(* IEC 61131-3 sources: JingjiangMoonbox/Application/Application/任务列表/Main_Task/套色调整/新算法/JIEOU, 8 files *)

(* ---- JIEOU10.st ---- *)
(*@CES
Name=JIEOU10
Type=FunctionBlock
TypeGuid=6f9dac99-8de1-4efc-8465-68ac443b7d08
Guid=2b28cbf0-4862-4f21-a282-23685e336d72
HasDeclaration=True
HasImplementation=True
*)
{DECLARATION}
FUNCTION JIEOU10 : REAL
VAR_INPUT
	i_rPI2_AND_JIEOU3_AND_JIEOU4:REAL;(*PI2和JIEOU3JIEOU4经过JIEOU8 Gc2Yk_K5_K6的输出/Gc2Uk_K5_K6输入*)
	i_rJIEOU5:REAL;(*U5经过JIEOU8 Gc2Yk_K3的输出/Gc2Uk_K4输入*)
	i_rJIEOU6:REAL;(*U6经过JIEOU9 Gc2Yk_K3的输出*)
	i_rJIEOU7:REAL;(*U7经过JIEOU9 Gc2_1的输出*)
	i_rJIEOU8:REAL;(*U8输出*)
	i_rJIEOU9:REAL;(*U9输出*)
	i_rPI10:REAL;(*PI10输出*)

	i_prU10: POINTER TO REAL;(*解耦后控制器8输出*)

(*
	i_rL:REAL;(*版周长mm*)
	i_rV:REAL;(*运行速度m/min*)
*)
	i_rTs:REAL;(*2024.6.29.135040修改为了输入@s*)
	i_rA:REAL;(*系统参数A*)
(*Gc1_1寄存器*)
	i_prGc1_1_Uk:POINTER TO ARRAY [1..ARC_DELAY_N_MAX] OF REAL;(*Gc1_1输入寄存器*)
	i_prGc1_1_Gc1_Yk:POINTER TO ARRAY [1..2] OF REAL;(*Gc1_1 Gc1输出寄存器*)
(*Gc2_1寄存器*)
	i_prGc2_1_Uk:POINTER TO ARRAY [1..ARC_DELAY_N_MAX] OF REAL;(*Gc2_1输入寄存器*)
	i_prGc2_1_Yk:POINTER TO ARRAY [1..2] OF REAL;(*Gc2_1输出寄存器*)

	i_prGc2_1_Gc1_Uk:POINTER TO ARRAY [1..2] OF REAL;(*Gc2_1 Gc1输入寄存器*)
	i_prGc2_1_Gc2_Yk:POINTER TO ARRAY [1..2] OF REAL;(*Gc2_1 Gc2输出寄存器*)

(*Gc2寄存器3*)
	i_prGc2Uk_K5:POINTER TO ARRAY [1..2] OF REAL;(*Gc2输入寄存器2*)
	i_prGc2Yk_K5:POINTER TO ARRAY [1..2] OF REAL;(*Gc2输出寄存器2*)

(*Gc2寄存器1*)
	i_prGc2Uk_K4:POINTER TO ARRAY [1..2] OF REAL;(*Gc2输入寄存器1*)
	i_prGc2Yk_K4:POINTER TO ARRAY [1..2] OF REAL;(*Gc2输出寄存器1*)
(*Gc2寄存器2*)
	i_prGc2Uk_K3:POINTER TO ARRAY [1..2] OF REAL;(*Gc2输入寄存器2*)
	i_prGc2Yk_K3:POINTER TO ARRAY [1..2] OF REAL;(*Gc2输出寄存器2*)

(*控制参数*)
	i_iN:INT;(*时延拍数N=TL/Ts+1*)
	i_bEn:BOOL;(*解耦使能 1：开解耦*)
	i_bK3:BOOL;(*K3=1时前三解耦*)
	i_bK4:BOOL;(*K4=1时前四解耦*)
	i_bK5:BOOL;(*K5=1时前五解耦*)
	i_bK6:BOOL;(*K6=1时前六解耦*)
END_VAR
VAR
(*	rTs:REAL:=0;(*采样时间*)   *)
	iI: INT:=0;

	(*中间变量*)
	rTemp5:REAL:=0;(*Gc2_K5输入*)
	rTemp6:REAL:=0;(*Gc2_K5输出*)

	rTemp7:REAL:=0;(*PI2+JIEOU3+JIEOU4输出*)

	(*中间变量*)
	rTemp1:REAL:=0;(*Gc2_K4输入*)
	rTemp2:REAL:=0;(*Gc2_K4输出*)
	(*中间变量*)
	rTemp3:REAL:=0;(*Gc2_K3输入*)
	rTemp4:REAL:=0;(*Gc2_K3输出*)

	rTempz:REAL:=0;(*总输出*)
	rGc1_1Out:REAL:=0;(*rGcd1_1控制器输出*)
	rGc2_1Out:REAL:=0;(*rGcd2_1控制器输出*)
END_VAR
{IMPLEMENTATION}
(*

(*更新寄存器*)

*)

(*计算*)
IF (i_bK5<>0 AND i_bK6<>0)  THEN
	rTemp5:=i_rPI2_AND_JIEOU3_AND_JIEOU4+i_rJIEOU5;
ELSIF (i_bK5<>0 AND i_bK6=0) THEN
	rTemp5:=i_rJIEOU5;
ELSE
	rTemp5:=0;
END_IF

Gc2(rTemp5,ADR(rTemp6),i_rTs,i_rA,i_prGc2Uk_K5,i_prGc2Yk_K5);
rTemp7:=rTemp6+i_rJIEOU6;

rTemp3:=i_rJIEOU7;
rTemp1:=rTemp7;
Gc2(rTemp1,ADR(rTemp2),i_rTs,i_rA,i_prGc2Uk_K4,i_prGc2Yk_K4);
Gc2(rTemp3,ADR(rTemp4),i_rTs,i_rA,i_prGc2Uk_K3,i_prGc2Yk_K3);

IF i_bK4=0 THEN
	rTemp2:=0;
	i_prGc2Yk_K4^[1]:=rTemp2;
END_IF

IF i_bK3=0 THEN
	rTemp4:=0;
	i_prGc2Yk_K3^[1]:=rTemp4;
END_IF

Gcd1_1(i_rJIEOU9,ADR(rGc1_1Out),i_rTs,i_rA,i_prGc1_1_Uk,i_prGc1_1_Gc1_Yk,i_iN,i_bEn);

Gcd2_1(i_rJIEOU8,ADR(rGc2_1Out),i_rTs,i_rA,i_prGc2_1_Uk,i_prGc2_1_Yk,i_prGc2_1_Gc1_Uk,i_prGc2_1_Gc2_Yk,i_iN,i_bEn);

rTempz:=rGc1_1Out+rGc2_1Out+i_rPI10+rTemp2+rTemp4;

(*输出*)
IF i_bEn<>0 THEN
	i_prU10^:=rTempz;
ELSE
	i_prU10^:=i_rPI10;
END_IF

(* ---- JIEOU3.st ---- *)
(*@CES
Name=JIEOU3
Type=FunctionBlock
TypeGuid=6f9dac99-8de1-4efc-8465-68ac443b7d08
Guid=7be6ac6f-cc63-4b01-8a46-0da4dcccc2cf
HasDeclaration=True
HasImplementation=True
*)
{DECLARATION}
FUNCTION JIEOU3 : REAL
VAR_INPUT

	i_rPI2:REAL;(*PI2输出*)
	i_rPI3:REAL;(*PI3输出*)

	i_prU3: POINTER TO REAL;(*解耦后控制器3输出*)

(*
	i_rL:REAL;(*版周长mm*)
	i_rV:REAL;(*运行速度m/min*)
*)
	i_rTs:REAL;(*2024.6.29.135040修改为了输入@s*)
	i_rA:REAL;(*系统参数A*)

	i_prGc1_1_Uk:POINTER TO ARRAY [1..ARC_DELAY_N_MAX] OF REAL;(*Gc1_1输入寄存器*)
	i_prGc1_1_Gc1_Yk:POINTER TO ARRAY [1..2] OF REAL;(*Gc1_1 Gc1输出寄存器*)

	i_iN:INT;(*时延拍数N=TL/Ts+1*)
	i_bEn:BOOL;(*解耦使能 1：开解耦*)
END_VAR

VAR
(*	rTs:REAL:=0;(*采样时间*)   *)

	iI: INT:=0;

	(*中间变量*)
	rTemp1:REAL:=0;(*总输出*)
	rGc1_1Out:REAL:=0;(*rGcd1_1控制器输出*)
END_VAR
{IMPLEMENTATION}
(*
(*更新寄存器*)
i_prGc1_1_Gc1_Yk^[2]:=i_prGc1_1_Gc1_Yk^[1];

FOR iI:=0 TO i_iN-2 BY 1 DO
	i_prGc1_1_Uk^[i_iN-iI]:=i_prGc1_1_Uk^[i_iN-iI-1];
END_FOR
*)

(*计算*)
Gcd1_1(i_rPI2,ADR(rGc1_1Out),i_rTs,i_rA,i_prGc1_1_Uk,i_prGc1_1_Gc1_Yk,i_iN,i_bEn);
rTemp1:=rGc1_1Out+i_rPI3;

(*输出*)
IF i_bEn<>0 THEN
	i_prU3^:=rTemp1;
ELSE
	i_prU3^:=i_rPI3;
END_IF

(* ---- JIEOU4.st ---- *)
(*@CES
Name=JIEOU4
Type=FunctionBlock
TypeGuid=6f9dac99-8de1-4efc-8465-68ac443b7d08
Guid=1946c078-7c38-40e6-bd29-bc69214024d3
HasDeclaration=True
HasImplementation=True
*)
{DECLARATION}
FUNCTION JIEOU4 : REAL
VAR_INPUT

	i_rPI2:REAL;(*PI2输出*)
	i_rJIEOU3:REAL;(*U3输出*)
	i_rPI4:REAL;(*PI4输出*)

	i_prU4: POINTER TO REAL;(*解耦后控制器4输出*)

(*
	i_rL:REAL;(*版周长mm*)
	i_rV:REAL;(*运行速度m/min*)
*)
	i_rTs:REAL;(*2024.6.29.135040修改为了输入@s*)
	i_rA:REAL;(*系统参数A*)
(*Gc1_1寄存器*)
	i_prGc1_1_Uk:POINTER TO ARRAY [1..ARC_DELAY_N_MAX] OF REAL;(*Gc1_1输入寄存器*)
	i_prGc1_1_Gc1_Yk:POINTER TO ARRAY [1..2] OF REAL;(*Gc1_1 Gc1输出寄存器*)
(*Gc2_1寄存器*)
	i_prGc2_1_Uk:POINTER TO ARRAY [1..ARC_DELAY_N_MAX] OF REAL;(*Gc2_1输入寄存器*)
	i_prGc2_1_Yk:POINTER TO ARRAY [1..2] OF REAL;(*Gc2_1输出寄存器*)

	i_prGc2_1_Gc1_Uk:POINTER TO ARRAY [1..2] OF REAL;(*Gc2_1 Gc1输入寄存器*)
	i_prGc2_1_Gc2_Yk:POINTER TO ARRAY [1..2] OF REAL;(*Gc2_1 Gc2输出寄存器*)

	i_iN:INT;(*时延拍数N=TL/Ts+1*)
	i_bEn:BOOL;(*解耦使能 1：开解耦*)
END_VAR

VAR
(*	rTs:REAL:=0;(*采样时间*)   *)
	iI: INT:=0;

	(*中间变量*)
	rTemp1:REAL:=0;(*总输出*)
	rGc1_1Out:REAL:=0;(*rGcd1_1控制器输出*)
	rGc2_1Out:REAL:=0;(*rGcd2_1控制器输出*)
END_VAR
{IMPLEMENTATION}
(*
(*更新寄存器*)
(*Gc1_1*)
i_prGc1_1_Gc1_Yk^[2]:=i_prGc1_1_Gc1_Yk^[1];

FOR iI:=0 TO i_iN-2 BY 1 DO
	i_prGc1_1_Uk^[i_iN-iI]:=i_prGc1_1_Uk^[i_iN-iI-1];
END_FOR

(*Gc2_1*)
i_prGc2_1_Gc1_Uk^[2]:=i_prGc2_1_Gc1_Uk^[1];

i_prGc2_1_Gc2_Yk^[2]:=i_prGc2_1_Gc2_Yk^[1];

i_prGc2_1_Yk^[2]:=i_prGc2_1_Yk^[1];

FOR iI:=0 TO i_iN-2 BY 1 DO
	i_prGc2_1_Uk^[i_iN-iI]:=i_prGc2_1_Uk^[i_iN-iI-1];
END_FOR
*)

(*计算*)
Gcd1_1(i_rJIEOU3,ADR(rGc1_1Out),i_rTs,i_rA,i_prGc1_1_Uk,i_prGc1_1_Gc1_Yk,i_iN,i_bEn);
Gcd2_1(i_rPI2,ADR(rGc2_1Out),i_rTs,i_rA,i_prGc2_1_Uk,i_prGc2_1_Yk,i_prGc2_1_Gc1_Uk,i_prGc2_1_Gc2_Yk,i_iN,i_bEn);
rTemp1:=rGc1_1Out+i_rPI4+rGc2_1Out;

(*输出*)
IF i_bEn<>0 THEN
	i_prU4^:=rTemp1;
ELSE
	i_prU4^:=i_rPI4;
END_IF

(* ---- JIEOU5.st ---- *)
(*@CES
Name=JIEOU5
Type=FunctionBlock
TypeGuid=6f9dac99-8de1-4efc-8465-68ac443b7d08
Guid=e0cca2d8-1a3c-4f43-93fd-67393267bfe9
HasDeclaration=True
HasImplementation=True
*)
{DECLARATION}
FUNCTION JIEOU5 : REAL
VAR_INPUT

	i_rPI2:REAL;(*PI2经过Gc2_1的输出*)
	i_rJIEOU3:REAL;(*U3输出*)
	i_rJIEOU4:REAL;(*U4输出*)
	i_rPI5:REAL;(*PI5输出*)

	i_prU5: POINTER TO REAL;(*解耦后控制器5输出*)

(*
	i_rL:REAL;(*版周长mm*)
	i_rV:REAL;(*运行速度m/min*)
*)
	i_rTs:REAL;(*2024.6.29.135040修改为了输入@s*)
	i_rA:REAL;(*系统参数A*)
(*Gc1_1寄存器*)
	i_prGc1_1_Uk:POINTER TO ARRAY [1..ARC_DELAY_N_MAX] OF REAL;(*Gc1_1输入寄存器*)
	i_prGc1_1_Gc1_Yk:POINTER TO ARRAY [1..2] OF REAL;(*Gc1_1 Gc1输出寄存器*)
(*Gc2_1寄存器*)
	i_prGc2_1_Uk:POINTER TO ARRAY [1..ARC_DELAY_N_MAX] OF REAL;(*Gc2_1输入寄存器*)
	i_prGc2_1_Yk:POINTER TO ARRAY [1..2] OF REAL;(*Gc2_1输出寄存器*)

	i_prGc2_1_Gc1_Uk:POINTER TO ARRAY [1..2] OF REAL;(*Gc2_1 Gc1输入寄存器*)
	i_prGc2_1_Gc2_Yk:POINTER TO ARRAY [1..2] OF REAL;(*Gc2_1 Gc2输出寄存器*)

(*Gc2寄存器1*)
	i_prGc2Uk_K3:POINTER TO ARRAY [1..2] OF REAL;(*Gc2输入寄存器1*)
	i_prGc2Yk_K3:POINTER TO ARRAY [1..2] OF REAL;(*Gc2输出寄存器1*)
(*控制参数*)
	i_iN:INT;(*时延拍数N=TL/Ts+1*)
	i_bEn:BOOL;(*解耦使能 1：开解耦*)
	i_bK3:BOOL;(*K3=1时前三解耦*)
END_VAR
VAR
(*	rTs:REAL:=0;(*采样时间*)   *)
	iI: INT:=0;

	(*中间变量*)
	rTemp1:REAL:=0;(*Gc2输入*)
	rTemp2:REAL:=0;(*Gc2输入*)

	rTempz:REAL:=0;(*总输出*)
	rGc1_1Out:REAL:=0;(*rGcd1_1控制器输出*)
	rGc2_1Out:REAL:=0;(*rGcd2_1控制器输出*)
END_VAR
{IMPLEMENTATION}
(*
(*更新寄存器*)

(*Gc1_1*)
i_prGc1_1_Gc1_Yk^[2]:=i_prGc1_1_Gc1_Yk^[1];

FOR iI:=0 TO i_iN-2 BY 1 DO
	i_prGc1_1_Uk^[i_iN-iI]:=i_prGc1_1_Uk^[i_iN-iI-1];
END_FOR

(*Gc2_1*)
i_prGc2_1_Gc1_Uk^[2]:=i_prGc2_1_Gc1_Uk^[1];

i_prGc2_1_Gc2_Yk^[2]:=i_prGc2_1_Gc2_Yk^[1];

i_prGc2_1_Yk^[2]:=i_prGc2_1_Yk^[1];

FOR iI:=0 TO i_iN-2 BY 1 DO
	i_prGc2_1_Uk^[i_iN-iI]:=i_prGc2_1_Uk^[i_iN-iI-1];
END_FOR

(*Gc2*)
i_prGc2Uk^[2]:=i_prGc2Uk^[1];
i_prGc2Yk^[2]:=i_prGc2Yk^[1];

*)

(*计算*)

rTemp1:=i_rPI2;
Gc2(rTemp1,ADR(rTemp2),i_rTs,i_rA,i_prGc2Uk_K3,i_prGc2Yk_K3);
IF i_bK3=0 THEN
	rTemp2:=0;
	i_prGc2Yk_K3^[1]:=rTemp2;
END_IF

Gcd1_1(i_rJIEOU4,ADR(rGc1_1Out),i_rTs,i_rA,i_prGc1_1_Uk,i_prGc1_1_Gc1_Yk,i_iN,i_bEn);

Gcd2_1(i_rJIEOU3,ADR(rGc2_1Out),i_rTs,i_rA,i_prGc2_1_Uk,i_prGc2_1_Yk,i_prGc2_1_Gc1_Uk,i_prGc2_1_Gc2_Yk,i_iN,i_bEn);

rTempz:=rGc1_1Out+rGc2_1Out+i_rPI5+rTemp2;

(*输出*)

(*输出*)
IF i_bEn<>0 THEN
	i_prU5^:=rTempz;
ELSE
	i_prU5^:=i_rPI5;
END_IF

(* ---- JIEOU6.st ---- *)
(*@CES
Name=JIEOU6
Type=FunctionBlock
TypeGuid=6f9dac99-8de1-4efc-8465-68ac443b7d08
Guid=de83d922-2817-4817-9257-b6b26cc19807
HasDeclaration=True
HasImplementation=True
*)
{DECLARATION}
FUNCTION JIEOU6 : REAL
VAR_INPUT
	i_rPI2:REAL;(*PI2经过JIEOU5_Gc2的输出/Gc2Uk_K4输入*)
	i_rJIEOU3:REAL;(*U3经过JIEOU5_Gcd2_1的输出/JIEOU3输出*)
	i_rJIEOU4:REAL;(*U4输出*)
	i_rJIEOU5:REAL;(*U5输出*)
	i_rPI6:REAL;(*PI6输出*)

	i_prU6: POINTER TO REAL;(*解耦后控制器6输出*)

(*
	i_rL:REAL;(*版周长mm*)
	i_rV:REAL;(*运行速度m/min*)
*)
	i_rTs:REAL;(*2024.6.29.135040修改为了输入@s*)
	i_rA:REAL;(*系统参数A*)
(*Gc1_1寄存器*)
	i_prGc1_1_Uk:POINTER TO ARRAY [1..ARC_DELAY_N_MAX] OF REAL;(*Gc1_1输入寄存器*)
	i_prGc1_1_Gc1_Yk:POINTER TO ARRAY [1..2] OF REAL;(*Gc1_1 Gc1输出寄存器*)
(*Gc2_1寄存器*)
	i_prGc2_1_Uk:POINTER TO ARRAY [1..ARC_DELAY_N_MAX] OF REAL;(*Gc2_1输入寄存器*)
	i_prGc2_1_Yk:POINTER TO ARRAY [1..2] OF REAL;(*Gc2_1输出寄存器*)

	i_prGc2_1_Gc1_Uk:POINTER TO ARRAY [1..2] OF REAL;(*Gc2_1 Gc1输入寄存器*)
	i_prGc2_1_Gc2_Yk:POINTER TO ARRAY [1..2] OF REAL;(*Gc2_1 Gc2输出寄存器*)

(*Gc2寄存器1*)
	i_prGc2Uk_K4:POINTER TO ARRAY [1..2] OF REAL;(*Gc2输入寄存器1*)
	i_prGc2Yk_K4:POINTER TO ARRAY [1..2] OF REAL;(*Gc2输出寄存器1*)
(*Gc2寄存器2*)
	i_prGc2Uk_K3:POINTER TO ARRAY [1..2] OF REAL;(*Gc2输入寄存器2*)
	i_prGc2Yk_K3:POINTER TO ARRAY [1..2] OF REAL;(*Gc2输出寄存器2*)
(*控制参数*)
	i_iN:INT;(*时延拍数N=TL/Ts+1*)
	i_bEn:BOOL;(*解耦使能 1：开解耦*)
	i_bK3:BOOL;(*K3=1时前三解耦*)
	i_bK4:BOOL;(*K4=1时前四解耦*)
END_VAR
VAR
(*	rTs:REAL:=0;(*采样时间*)   *)
	iI: INT:=0;

	(*中间变量*)
	rTemp1:REAL:=0;(*Gc2_K4输入*)
	rTemp2:REAL:=0;(*Gc2_K4输出*)
	(*中间变量*)
	rTemp3:REAL:=0;(*Gc2_K3输入*)
	rTemp4:REAL:=0;(*Gc2_K3输出*)

	rTempz:REAL:=0;(*总输出*)
	rGc1_1Out:REAL:=0;(*rGcd1_1控制器输出*)
	rGc2_1Out:REAL:=0;(*rGcd2_1控制器输出*)
END_VAR
{IMPLEMENTATION}
(*
(*更新寄存器*)

(*Gc1_1*)
i_prGc1_1_Gc1_Yk^[2]:=i_prGc1_1_Gc1_Yk^[1];

FOR iI:=0 TO i_iN-2 BY 1 DO
	i_prGc1_1_Uk^[i_iN-iI]:=i_prGc1_1_Uk^[i_iN-iI-1];
END_FOR

(*Gc2_1*)
i_prGc2_1_Gc1_Uk^[2]:=i_prGc2_1_Gc1_Uk^[1];

i_prGc2_1_Gc2_Yk^[2]:=i_prGc2_1_Gc2_Yk^[1];

i_prGc2_1_Yk^[2]:=i_prGc2_1_Yk^[1];

FOR iI:=0 TO i_iN-2 BY 1 DO
	i_prGc2_1_Uk^[i_iN-iI]:=i_prGc2_1_Uk^[i_iN-iI-1];
END_FOR

(*Gc2*)
i_prGc2Uk_K4^[2]:=i_prGc2Uk_K4^[1];
i_prGc2Yk_K4^[2]:=i_prGc2Yk_K4^[1];

(*Gc2*)
i_prGc2Uk_K3^[2]:=i_prGc2Uk_K3^[1];
i_prGc2Yk_K3^[2]:=i_prGc2Yk_K3^[1];
*)

(*计算*)
rTemp1:=i_rPI2;
rTemp3:=i_rJIEOU3;
Gc2(rTemp1,ADR(rTemp2),i_rTs,i_rA,i_prGc2Uk_K4,i_prGc2Yk_K4);
Gc2(rTemp3,ADR(rTemp4),i_rTs,i_rA,i_prGc2Uk_K3,i_prGc2Yk_K3);

IF i_bK4=0 THEN
	rTemp2:=0;
	i_prGc2Yk_K4^[1]:=rTemp2;
END_IF

IF i_bK3=0 THEN
	rTemp4:=0;
	i_prGc2Yk_K3^[1]:=rTemp4;
END_IF

Gcd1_1(i_rJIEOU5,ADR(rGc1_1Out),i_rTs,i_rA,i_prGc1_1_Uk,i_prGc1_1_Gc1_Yk,i_iN,i_bEn);

Gcd2_1(i_rJIEOU4,ADR(rGc2_1Out),i_rTs,i_rA,i_prGc2_1_Uk,i_prGc2_1_Yk,i_prGc2_1_Gc1_Uk,i_prGc2_1_Gc2_Yk,i_iN,i_bEn);

rTempz:=rGc1_1Out+rGc2_1Out+i_rPI6+rTemp2+rTemp4;

(*输出*)
IF i_bEn<>0 THEN
	i_prU6^:=rTempz;
ELSE
	i_prU6^:=i_rPI6;
END_IF

(* ---- JIEOU7.st ---- *)
(*@CES
Name=JIEOU7
Type=FunctionBlock
TypeGuid=6f9dac99-8de1-4efc-8465-68ac443b7d08
Guid=42a7d55e-0b4b-4417-9f25-6f09beff2d86
HasDeclaration=True
HasImplementation=True
*)
{DECLARATION}
FUNCTION JIEOU7 : REAL
VAR_INPUT
	i_rPI2:REAL;(*PI2经过JIEOU6_Gc2的输出/Gc2Uk_K5输入*)
	i_rJIEOU3:REAL;(*U3经过JIEOU6_Gcd2_1_G2的输出/JIEOU3输出*)
	i_rJIEOU4:REAL;(*U4输出/经过JIEOU6_Gcd2_1的输出*)
	i_rJIEOU5:REAL;(*U5输出*)
	i_rJIEOU6:REAL;(*U5输出*)
	i_rPI7:REAL;(*PI7输出*)

	i_prU7: POINTER TO REAL;(*解耦后控制器7输出*)

(*
	i_rL:REAL;(*版周长mm*)
	i_rV:REAL;(*运行速度m/min*)
*)
	i_rTs:REAL;(*2024.6.29.135040修改为了输入@s*)
	i_rA:REAL;(*系统参数A*)
(*Gc1_1寄存器*)
	i_prGc1_1_Uk:POINTER TO ARRAY [1..ARC_DELAY_N_MAX] OF REAL;(*Gc1_1输入寄存器*)
	i_prGc1_1_Gc1_Yk:POINTER TO ARRAY [1..2] OF REAL;(*Gc1_1 Gc1输出寄存器*)
(*Gc2_1寄存器*)
	i_prGc2_1_Uk:POINTER TO ARRAY [1..ARC_DELAY_N_MAX] OF REAL;(*Gc2_1输入寄存器*)
	i_prGc2_1_Yk:POINTER TO ARRAY [1..2] OF REAL;(*Gc2_1输出寄存器*)

	i_prGc2_1_Gc1_Uk:POINTER TO ARRAY [1..2] OF REAL;(*Gc2_1 Gc1输入寄存器*)
	i_prGc2_1_Gc2_Yk:POINTER TO ARRAY [1..2] OF REAL;(*Gc2_1 Gc2输出寄存器*)

(*Gc2寄存器1*)
	i_prGc2Uk_K4:POINTER TO ARRAY [1..2] OF REAL;(*Gc2输入寄存器1*)
	i_prGc2Yk_K4:POINTER TO ARRAY [1..2] OF REAL;(*Gc2输出寄存器1*)
(*Gc2寄存器2*)
	i_prGc2Uk_K3:POINTER TO ARRAY [1..2] OF REAL;(*Gc2输入寄存器2*)
	i_prGc2Yk_K3:POINTER TO ARRAY [1..2] OF REAL;(*Gc2输出寄存器2*)
(*控制参数*)
	i_iN:INT;(*时延拍数N=TL/Ts+1*)
	i_bEn:BOOL;(*解耦使能 1：开解耦*)
	i_bK3:BOOL;(*K3=1时前三解耦*)
	i_bK4:BOOL;(*K4=1时前四解耦*)
	i_bK5:BOOL;(*K5=1时前五解耦*)
END_VAR
VAR
(*	rTs:REAL:=0;(*采样时间*)   *)
	iI: INT:=0;

	(*中间变量*)
	rTemp1:REAL:=0;(*Gc2_K4输入*)
	rTemp2:REAL:=0;(*Gc2_K4输出*)
	(*中间变量*)
	rTemp3:REAL:=0;(*Gc2_K3输入*)
	rTemp4:REAL:=0;(*Gc2_K3输出*)

	rTempz:REAL:=0;(*总输出*)
	rGc1_1Out:REAL:=0;(*rGcd1_1控制器输出*)
	rGc2_1Out:REAL:=0;(*rGcd2_1控制器输出*)
END_VAR
{IMPLEMENTATION}
(*
(*更新寄存器*)

(*Gc1_1*)
i_prGc1_1_Gc1_Yk^[2]:=i_prGc1_1_Gc1_Yk^[1];

FOR iI:=0 TO i_iN-2 BY 1 DO
	i_prGc1_1_Uk^[i_iN-iI]:=i_prGc1_1_Uk^[i_iN-iI-1];
END_FOR

(*Gc2_1*)
i_prGc2_1_Gc1_Uk^[2]:=i_prGc2_1_Gc1_Uk^[1];

i_prGc2_1_Gc2_Yk^[2]:=i_prGc2_1_Gc2_Yk^[1];

i_prGc2_1_Yk^[2]:=i_prGc2_1_Yk^[1];

FOR iI:=0 TO i_iN-2 BY 1 DO
	i_prGc2_1_Uk^[i_iN-iI]:=i_prGc2_1_Uk^[i_iN-iI-1];
END_FOR

(*Gc2*)
i_prGc2Uk_K4^[2]:=i_prGc2Uk_K4^[1];
i_prGc2Yk_K4^[2]:=i_prGc2Yk_K4^[1];

(*Gc2*)
i_prGc2Uk_K3^[2]:=i_prGc2Uk_K3^[1];
i_prGc2Yk_K3^[2]:=i_prGc2Yk_K3^[1];
*)

(*计算*)
IF (i_bK5<>0 AND i_bK4<>0)  THEN
	rTemp1:=i_rPI2+i_rJIEOU3;
ELSIF (i_bK5=0 AND i_bK4<>0) THEN
	rTemp1:=i_rJIEOU3;
ELSE
	rTemp1:=0;
END_IF

Gc2(rTemp1,ADR(rTemp2),i_rTs,i_rA,i_prGc2Uk_K4,i_prGc2Yk_K4);

rTemp3:=i_rJIEOU4;
Gc2(rTemp3,ADR(rTemp4),i_rTs,i_rA,i_prGc2Uk_K3,i_prGc2Yk_K3);
IF i_bK3=0 THEN
	rTemp4:=0;
	i_prGc2Yk_K3^[1]:=rTemp4;
END_IF

Gcd1_1(i_rJIEOU6,ADR(rGc1_1Out),i_rTs,i_rA,i_prGc1_1_Uk,i_prGc1_1_Gc1_Yk,i_iN,i_bEn);

Gcd2_1(i_rJIEOU5,ADR(rGc2_1Out),i_rTs,i_rA,i_prGc2_1_Uk,i_prGc2_1_Yk,i_prGc2_1_Gc1_Uk,i_prGc2_1_Gc2_Yk,i_iN,i_bEn);

rTempz:=rGc1_1Out+rGc2_1Out+i_rPI7+rTemp2+rTemp4;

(*输出*)
IF i_bEn<>0 THEN
	i_prU7^:=rTempz;
ELSE
	i_prU7^:=i_rPI7;
END_IF

(* ---- JIEOU8.st ---- *)
(*@CES
Name=JIEOU8
Type=FunctionBlock
TypeGuid=6f9dac99-8de1-4efc-8465-68ac443b7d08
Guid=cb531a50-6479-4a30-ae73-c8a7aeed7012
HasDeclaration=True
HasImplementation=True
*)
{DECLARATION}
FUNCTION JIEOU8 : REAL
VAR_INPUT
	i_rPI2:REAL;(*PI2经过JIEOU6 Gc2Yk_K4的输出/Gc2Uk_K5_K6输入*)
	i_rJIEOU3:REAL;(*U3经过JIEOU6 Gc2Yk_K3的输出/Gc2Uk_K5输入*)
	i_rJIEOU4:REAL;(*U4经过JIEOU7 Gc2Yk_K3的输出*)
	i_rJIEOU5:REAL;(*U5经过JIEOU7 Gc2_1的输出*)
	i_rJIEOU6:REAL;(*U6输出*)
	i_rJIEOU7:REAL;(*U7输出*)
	i_rPI8:REAL;(*PI8输出*)

	i_prU8: POINTER TO REAL;(*解耦后控制器8输出*)

(*
	i_rL:REAL;(*版周长mm*)
	i_rV:REAL;(*运行速度m/min*)
*)
	i_rTs:REAL;(*2024.6.29.135040修改为了输入@s*)
	i_rA:REAL;(*系统参数A*)
(*Gc1_1寄存器*)
	i_prGc1_1_Uk:POINTER TO ARRAY [1..ARC_DELAY_N_MAX] OF REAL;(*Gc1_1输入寄存器*)
	i_prGc1_1_Gc1_Yk:POINTER TO ARRAY [1..2] OF REAL;(*Gc1_1 Gc1输出寄存器*)
(*Gc2_1寄存器*)
	i_prGc2_1_Uk:POINTER TO ARRAY [1..ARC_DELAY_N_MAX] OF REAL;(*Gc2_1输入寄存器*)
	i_prGc2_1_Yk:POINTER TO ARRAY [1..2] OF REAL;(*Gc2_1输出寄存器*)

	i_prGc2_1_Gc1_Uk:POINTER TO ARRAY [1..2] OF REAL;(*Gc2_1 Gc1输入寄存器*)
	i_prGc2_1_Gc2_Yk:POINTER TO ARRAY [1..2] OF REAL;(*Gc2_1 Gc2输出寄存器*)

(*Gc2寄存器3*)
	i_prGc2Uk_K5:POINTER TO ARRAY [1..2] OF REAL;(*Gc2输入寄存器2*)
	i_prGc2Yk_K5:POINTER TO ARRAY [1..2] OF REAL;(*Gc2输出寄存器2*)

(*Gc2寄存器1*)
	i_prGc2Uk_K4:POINTER TO ARRAY [1..2] OF REAL;(*Gc2输入寄存器1*)
	i_prGc2Yk_K4:POINTER TO ARRAY [1..2] OF REAL;(*Gc2输出寄存器1*)
(*Gc2寄存器2*)
	i_prGc2Uk_K3:POINTER TO ARRAY [1..2] OF REAL;(*Gc2输入寄存器2*)
	i_prGc2Yk_K3:POINTER TO ARRAY [1..2] OF REAL;(*Gc2输出寄存器2*)

(*控制参数*)
	i_iN:INT;(*时延拍数N=TL/Ts+1*)
	i_bEn:BOOL;(*解耦使能 1：开解耦*)
	i_bK3:BOOL;(*K3=1时前三解耦*)
	i_bK4:BOOL;(*K4=1时前四解耦*)
	i_bK5:BOOL;(*K5=1时前五解耦*)
	i_bK6:BOOL;(*K6=1时前六解耦*)
END_VAR
VAR
(*	rTs:REAL:=0;(*采样时间*)   *)
	iI: INT:=0;

	(*中间变量*)
	rTemp5:REAL:=0;(*Gc2_K5输入*)
	rTemp6:REAL:=0;(*Gc2_K5输出*)

	rTemp7:REAL:=0;(*PI2+JIEOU3+JIEOU4输出*)

	(*中间变量*)
	rTemp1:REAL:=0;(*Gc2_K4输入*)
	rTemp2:REAL:=0;(*Gc2_K4输出*)
	(*中间变量*)
	rTemp3:REAL:=0;(*Gc2_K3输入*)
	rTemp4:REAL:=0;(*Gc2_K3输出*)

	rTempz:REAL:=0;(*总输出*)
	rGc1_1Out:REAL:=0;(*rGcd1_1控制器输出*)
	rGc2_1Out:REAL:=0;(*rGcd2_1控制器输出*)
END_VAR
{IMPLEMENTATION}
Gc2(rTemp1,ADR(rTemp2),i_rTs,i_rA,i_prGc2Uk_K4,i_prGc2Yk_K4);
Gc2(rTemp3,ADR(rTemp4),i_rTs,i_rA,i_prGc2Uk_K3,i_prGc2Yk_K3);

IF i_bK4=0 THEN
	rTemp2:=0;
	i_prGc2Yk_K4^[1]:=rTemp2;
END_IF

IF i_bK3=0 THEN
	rTemp4:=0;
	i_prGc2Yk_K3^[1]:=rTemp4;
END_IF

Gcd1_1(i_rJIEOU7,ADR(rGc1_1Out),i_rTs,i_rA,i_prGc1_1_Uk,i_prGc1_1_Gc1_Yk,i_iN,i_bEn);

Gcd2_1(i_rJIEOU6,ADR(rGc2_1Out),i_rTs,i_rA,i_prGc2_1_Uk,i_prGc2_1_Yk,i_prGc2_1_Gc1_Uk,i_prGc2_1_Gc2_Yk,i_iN,i_bEn);

rTempz:=rGc1_1Out+rGc2_1Out+i_rPI8+rTemp2+rTemp4;

(*输出*)
IF i_bEn<>0 THEN
	i_prU8^:=rTempz;
ELSE
	i_prU8^:=i_rPI8;
END_IF

(* ---- JIEOU9.st ---- *)
(*@CES
Name=JIEOU9
Type=FunctionBlock
TypeGuid=6f9dac99-8de1-4efc-8465-68ac443b7d08
Guid=4b016c4b-4091-44a0-b80a-ccae90087a29
HasDeclaration=True
HasImplementation=True
*)
{DECLARATION}
FUNCTION JIEOU9 : REAL
VAR_INPUT
	i_rPI2:REAL;(*PI2经过JIEOU6 Gc2Yk_K4的输出/Gc2Uk_K5_K6输入*)
	i_rJIEOU3:REAL;(*U3经过JIEOU6 Gc2Yk_K3的输出/Gc2Uk_K5输入*)
	i_rJIEOU4:REAL;(*U4经过JIEOU7 Gc2Yk_K3的输出*)
	i_rJIEOU5:REAL;(*U5经过JIEOU7 Gc2_1的输出*)
	i_rJIEOU6:REAL;(*U6输出*)
	i_rJIEOU7:REAL;(*U7输出*)
	i_rPI8:REAL;(*PI8输出*)

	i_prU8: POINTER TO REAL;(*解耦后控制器8输出*)

(*
	i_rL:REAL;(*版周长mm*)
	i_rV:REAL;(*运行速度m/min*)
*)
	i_rTs:REAL;(*2024.6.29.135040修改为了输入@s*)
	i_rA:REAL;(*系统参数A*)
(*Gc1_1寄存器*)
	i_prGc1_1_Uk:POINTER TO ARRAY [1..ARC_DELAY_N_MAX] OF REAL;(*Gc1_1输入寄存器*)
	i_prGc1_1_Gc1_Yk:POINTER TO ARRAY [1..2] OF REAL;(*Gc1_1 Gc1输出寄存器*)
(*Gc2_1寄存器*)
	i_prGc2_1_Uk:POINTER TO ARRAY [1..ARC_DELAY_N_MAX] OF REAL;(*Gc2_1输入寄存器*)
	i_prGc2_1_Yk:POINTER TO ARRAY [1..2] OF REAL;(*Gc2_1输出寄存器*)

	i_prGc2_1_Gc1_Uk:POINTER TO ARRAY [1..2] OF REAL;(*Gc2_1 Gc1输入寄存器*)
	i_prGc2_1_Gc2_Yk:POINTER TO ARRAY [1..2] OF REAL;(*Gc2_1 Gc2输出寄存器*)

(*Gc2寄存器3*)
	i_prGc2Uk_K5:POINTER TO ARRAY [1..2] OF REAL;(*Gc2输入寄存器2*)
	i_prGc2Yk_K5:POINTER TO ARRAY [1..2] OF REAL;(*Gc2输出寄存器2*)

(*Gc2寄存器1*)
	i_prGc2Uk_K4:POINTER TO ARRAY [1..2] OF REAL;(*Gc2输入寄存器1*)
	i_prGc2Yk_K4:POINTER TO ARRAY [1..2] OF REAL;(*Gc2输出寄存器1*)
(*Gc2寄存器2*)
	i_prGc2Uk_K3:POINTER TO ARRAY [1..2] OF REAL;(*Gc2输入寄存器2*)
	i_prGc2Yk_K3:POINTER TO ARRAY [1..2] OF REAL;(*Gc2输出寄存器2*)

(*控制参数*)
	i_iN:INT;(*时延拍数N=TL/Ts+1*)
	i_bEn:BOOL;(*解耦使能 1：开解耦*)
	i_bK3:BOOL;(*K3=1时前三解耦*)
	i_bK4:BOOL;(*K4=1时前四解耦*)
	i_bK5:BOOL;(*K5=1时前五解耦*)
	i_bK6:BOOL;(*K6=1时前六解耦*)
END_VAR
VAR
(*	rTs:REAL:=0;(*采样时间*)   *)
	iI: INT:=0;

	(*中间变量*)
	rTemp5:REAL:=0;(*Gc2_K5输入*)
	rTemp6:REAL:=0;(*Gc2_K5输出*)

	rTemp7:REAL:=0;(*PI2+JIEOU3+JIEOU4输出*)

	(*中间变量*)
	rTemp1:REAL:=0;(*Gc2_K4输入*)
	rTemp2:REAL:=0;(*Gc2_K4输出*)
	(*中间变量*)
	rTemp3:REAL:=0;(*Gc2_K3输入*)
	rTemp4:REAL:=0;(*Gc2_K3输出*)

	rTempz:REAL:=0;(*总输出*)
	rGc1_1Out:REAL:=0;(*rGcd1_1控制器输出*)
	rGc2_1Out:REAL:=0;(*rGcd2_1控制器输出*)
END_VAR
{IMPLEMENTATION}
(*
(*更新寄存器*)

(*Gc1_1*)
i_prGc1_1_Gc1_Yk^[2]:=i_prGc1_1_Gc1_Yk^[1];

FOR iI:=0 TO i_iN-2 BY 1 DO
	i_prGc1_1_Uk^[i_iN-iI]:=i_prGc1_1_Uk^[i_iN-iI-1];
END_FOR

(*Gc2_1*)
i_prGc2_1_Gc1_Uk^[2]:=i_prGc2_1_Gc1_Uk^[1];

i_prGc2_1_Gc2_Yk^[2]:=i_prGc2_1_Gc2_Yk^[1];

i_prGc2_1_Yk^[2]:=i_prGc2_1_Yk^[1];

FOR iI:=0 TO i_iN-2 BY 1 DO
	i_prGc2_1_Uk^[i_iN-iI]:=i_prGc2_1_Uk^[i_iN-iI-1];
END_FOR

(*Gc2*)
i_prGc2Uk_K5^[2]:=i_prGc2Uk_K5^[1];
i_prGc2Yk_K5^[2]:=i_prGc2Yk_K5^[1];

(*Gc2*)
i_prGc2Uk_K4^[2]:=i_prGc2Uk_K4^[1];
i_prGc2Yk_K4^[2]:=i_prGc2Yk_K4^[1];

(*Gc2*)
i_prGc2Uk_K3^[2]:=i_prGc2Uk_K3^[1];
i_prGc2Yk_K3^[2]:=i_prGc2Yk_K3^[1];
*)

(*计算*)
IF (i_bK5<>0 AND i_bK6<>0)  THEN
	rTemp5:=i_rPI2+i_rJIEOU3;
ELSIF (i_bK5<>0 AND i_bK6=0) THEN
	rTemp5:=i_rJIEOU3;
ELSE
	rTemp5:=0;
END_IF

Gc2(rTemp5,ADR(rTemp6),i_rTs,i_rA,i_prGc2Uk_K5,i_prGc2Yk_K5);
rTemp7:=rTemp6+i_rJIEOU4;

rTemp3:=i_rJIEOU5;
rTemp1:=rTemp7;
Gc2(rTemp1,ADR(rTemp2),i_rTs,i_rA,i_prGc2Uk_K4,i_prGc2Yk_K4);
Gc2(rTemp3,ADR(rTemp4),i_rTs,i_rA,i_prGc2Uk_K3,i_prGc2Yk_K3);

IF i_bK4=0 THEN
	rTemp2:=0;
	i_prGc2Yk_K4^[1]:=rTemp2;
END_IF

IF i_bK3=0 THEN
	rTemp4:=0;
	i_prGc2Yk_K3^[1]:=rTemp4;
END_IF

Gcd1_1(i_rJIEOU7,ADR(rGc1_1Out),i_rTs,i_rA,i_prGc1_1_Uk,i_prGc1_1_Gc1_Yk,i_iN,i_bEn);

Gcd2_1(i_rJIEOU6,ADR(rGc2_1Out),i_rTs,i_rA,i_prGc2_1_Uk,i_prGc2_1_Yk,i_prGc2_1_Gc1_Uk,i_prGc2_1_Gc2_Yk,i_iN,i_bEn);

rTempz:=rGc1_1Out+rGc2_1Out+i_rPI8+rTemp2+rTemp4;

(*输出*)
IF i_bEn<>0 THEN
	i_prU8^:=rTempz;
ELSE
	i_prU8^:=i_rPI8;
END_IF
